// TIA Portal V21 export
// export: Created 2026-10-23T21:22:23.0525591Z, ExportSetting WithReadOnly, DisplayName Totally Integrated Automation Portal, DisplayVersion V21 Update 1, DisplayName SINAMICS Startdrive Advanced, DisplayVersion V21 HF2, DisplayName SINAMICS Startdrive G110M, G120, G120C, G120D, G120P, G115D, DisplayVersion V21 HF2, DisplayName SINAMICS Startdrive G130, G150, S120, S150, G200, G220, S200, S210, S220, Innomotics MVD, DisplayVersion V21 HF2, DisplayName STEP 7 Professional, DisplayVersion V21 Update 1, DisplayName STEP 7 Safety, DisplayVersion V21, DisplayName Tech WebApplication, DisplayVersion V21, DisplayName WinCC Basic/Comfort/Advanced, DisplayVersion V21 Update 1, DisplayName WinCC Unified, DisplayVersion V21 Update 1
ORGANIZATION_BLOCK "OB_DiagError"   // OB82, SCL, DiagnosticErrorInterrupt
TITLE = Diagnosefehleralarm / Diagnostic error interrupt
{ S7_Optimized_Access := 'TRUE' }
// Minimaler Diagnosefehler-OB / Minimal diagnostic error OB
// stored: CodeModifiedDate 2026-10-23T19:38:39.0176487Z, CompileDate 2026-10-23T19:38:39.0176487Z, ConstantName OB_OB_DiagError, CreationDate 2026-10-23T19:37:59.6610761Z, DownloadDate 0001-01-01T00:00:00Z, EventClass Diagnostic interrupt, InterfaceModifiedDate 2008-07-22T16:55:41.2736645Z, IsConsistent true, LoadMemoryLength 3699, ModifiedDate 2026-10-23T19:38:39.0176487Z, ParameterModified 2008-07-22T16:55:41.2736645Z, PriorityNumber 7, ProcessImagePartNumber 65535, SetENOAutomatically false, StructureModified 2008-07-22T16:55:41.2736645Z, WorkMemoryLength 120
   VAR_INPUT
      IO_State : Word;   // IO state of the HW object
      LADDR : HW_ANY;   // Hardware identifier
      Channel : UInt;   // Channel number
      MultiError : Bool;   // =true if more than one error is present
   END_VAR
BEGIN

       // Flag the diagnostic event
       "DB_Machine".StatusWord := "DB_Machine".StatusWord OR 16#0001;
END_ORGANIZATION_BLOCK
